Fanuc TP program (LS listing): SubProg2.LS

/PROG  SubProg2
/ATTR
OWNER		= MNEDITOR;
COMMENT		= "RoboDK sequence";
PROG_SIZE	= 0;
CREATE		= DATE 31-12-14  TIME 12:00:00;
MODIFIED	= DATE 31-12-14  TIME 12:00:00;
FILE_NAME	= SubProg2;
VERSION		= 0;
LINE_COUNT	= 1;
MEMORY_SIZE	= 0;
PROTECT		= READ_WRITE;
TCD:  STACK_SIZE	= 0,
      TASK_PRIORITY	= 50,
      TIME_SLICE	= 0,
      BUSY_LAMP_OFF	= 0,
      ABORT_REQUEST	= 0,
      PAUSE_REQUEST	= 0;
DEFAULT_GROUP	= 1,*,*,*,*,*,*;
CONTROL_CODE	= 00000000 00000000;
/MN
   1:J P[1] 20% FINE ;
/POS
P[1]{
   GP1:
    UF : 9, UT : 9,
	J1=    20.000 deg,	J2=    -10.000 deg,	J3=    20.000 deg,
	J4=    0.000 deg,	J5=    30.000 deg,	J6=    0.000 deg
};
/END
